// TIA Portal V19 export
TYPE "EM_Interface"
   STRUCT
      Cmds : Struct   // Comandos
         ManMode : Bool;   // Modo manual
         AutoMode : Bool;   // Modo automatico
         MaintenanceMode : Bool;   // Modo de mantenimiento
         Task : UInt;   // Codigo de tarea
         Execute : Bool;   // Ejecutar
         Reset : Bool;   // Reiniciar
         Hold : Bool;   // Retener
      END_STRUCT;
      Status : Struct   // Estado del EM
         ActiveTask : UInt;   // Tarea activa
         Ready : Bool;
         Busy : Bool;
         Done : Bool;
         Held : Bool;
         Error : Bool;
         ErrorID : UInt;
         AutAct : Bool;
         ManAct : Bool;
         Maintenance : Bool;
      END_STRUCT;
      Params : Struct   // Parametros
         ParamsReal : Array[0..8] of Real;
         ParamsInt : Array[0..8] of Int;
         ParamsBool : Array[0..8] of Bool;
      END_STRUCT;
   END_STRUCT;
END_TYPE
